// TIA Portal V20 export
FUNCTION_BLOCK "08_Systemzeit"   // FB167, LAD
{ S7_Optimized_Access := 'TRUE' }
// stored: MemoryReserve 100, SetENOAutomatically false
   VAR
      outputTIME : Date_And_Time;
      returnValue : Int;
      inputTIME : Date_And_Time;
      returnValueT : Int;
      execute : Bool;
   END_VAR
BEGIN

REGION Network 1: Aktuelles Datum und Uhrzeit auslesen
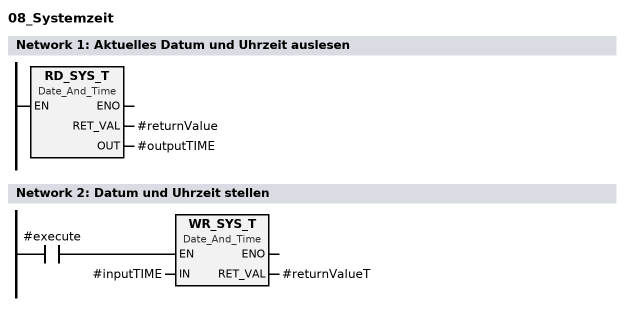
   RUNG wire#powerrail
      { S7_Templates := "date_type := Date_And_Time" } RD_SYS_T(RET_VAL => #returnValue, OUT => #outputTIME)
   END_RUNG
   // the same network as SCL:
   #returnValue := RD_SYS_T(OUT => #outputTIME);
END_REGION

REGION Network 2: Datum und Uhrzeit stellen
   RUNG wire#powerrail
      Contact( #execute )
      { S7_Templates := "date_type := Date_And_Time" } WR_SYS_T(IN := #inputTIME, RET_VAL => #returnValueT)
   END_RUNG
   // the same network as SCL:
   IF #execute THEN #returnValueT := WR_SYS_T(IN := #inputTIME); END_IF;
END_REGION
END_FUNCTION_BLOCK
